// TIA Portal V21 export
TagTable "T_V9"
  Y_V9 :   (PLC tag HMI_IF.BtnInit, HMI_Connection_1)
